TYPE E_ControlMode :
(
    IDLE        := 0,
    POSITION    := 1,
    VELOCITY    := 2,
    TORQUE      := 3
) UDINT := IDLE;
END_TYPE

(* stored: Version 1.1.0.1, ProductVersion 3.1.4026.18
   DUT E_ControlMode: Id {3fc01c8a-0e04-406b-aae4-37d5a08c513e} *)
